(* IEC 61131-3 sources: Lasal-MCP/examples/SampleSource/LASALScreenAdvancedSolution/LASALScreenAdvancedSolution/LASALScreenAdvacnedSolution/Stations/Terminal/HMI/Class/MyFirstMyIO, 1 file *)

(* ---- MyFirstMyIO.st ---- *)
(*!
<Class
	Name               = "MyFirstMyIO"
	Revision           = "0.0"
	RealtimeTask       = "false"
	CyclicTask         = "false"
	BackgroundTask     = "false"
	Sigmatek           = "false"
	OSInterface        = "false"
	HighPriority       = "false"
	Automatic          = "false"
	UpdateMode         = "Prescan"
	SharedCommandTable = "true"
	Objectsize         = "(450,180)">
	<Channels>
		<Server Name="Number" Visualized="false" Initialize="false" WriteProtected="true" Retentive="false"/>
		<Client Name="_Grafix" Required="false" Internal="false"/>
	</Channels>
	<Network Name="MyFirstMyIO">
		<!-- List of Components in this network -->
		<Components>
			<Object
				Name       = "_base"
				Class      = "_MyIO"
				Position   = "(218,120)"
				Visualized = "true"
				Remotely   = "true">
				<Channels>
					<Server Name="Refresh"/>
					<Server Name="Server0"/>
					<Client Name="Graphic"/>
					<Client Name="Lse"/>
				</Channels>
			</Object>
		</Components>
		<Comments>
		</Comments>
		<!-- List of Connections in this network -->
		<Connections>
			<Connection Source="this.Server0" Destination="_base.Server0" Vertices="(706,210),(534,210),"/>
			<Connection Source="this.Refresh" Destination="_base.Refresh" Vertices="(706,270),(534,270),"/>
			<Connection Source="_base.Lse" Destination="this.Lse" Vertices="(218,210),(38,210),"/>
		</Connections>
		<!-- Headerfiles -->
		<Options>
		</Options>
	</Network>
</Class>
*)
#pragma using _MyIO

MyFirstMyIO : CLASS
: _MyIO
  //Servers:
	Number 	: SvrCh_DINT;
  //Clients:
	_Grafix 	: CltChCmd__Grafix;
  //Variables:
  //Functions:
				//! <Function Comment="this method is called everytime when system wants to redraw the io" Name="Draw"/>
	FUNCTION __CDECL VIRTUAL GLOBAL Draw
		VAR_INPUT
			pio 	: ^_IO;			//! <Variable Comment="pointer to _IO information" Name="Draw.pio"/>
			pr 	: ^_RESULT;			//! <Variable Comment="pointer to _RESULT information" Name="Draw.pr"/>
			pv 	: ^_VARIABLE;			//! <Variable Comment="pointer to io _VARIABLE information" Name="Draw.pv"/>
			input 	: BOOL;			//! <Variable Comment="TRUE it&apos;s an input&#13;&#10;FALSE it&apos;s an output" Name="Draw.input"/>
		END_VAR
		VAR_OUTPUT
			retcode (EAX) 	: _DOIT;			//! <Variable Comment="for the returnstatement there are 3 different possibilities&#13;&#10;  _IDLE ..... the system should goon like it is (system goes on)&#13;&#10;  _IDIDIT ... i did it (system is ready)&#13;&#10;  _IFAILED .. i tried to do my best, but i failed (system is re" Name="Draw.retcode"/>
		END_VAR;
				//! <Function Comment="method is called cyclic during object is on screen&#13;&#10;&#13;&#10;pio ....... &#13;&#10;input .... TRUE it&apos;s an input / FALSE it&apos;s an output&#13;&#10;" Name="IF_Run"/>
	FUNCTION __CDECL VIRTUAL GLOBAL IF_Run
		VAR_INPUT
			pio 	: ^_IO;			//! <Variable Comment="pointer to _IO information given by LSE" Name="IF_Run.pio"/>
			input 	: BOOL;			//! <Variable Comment="TRUE it&apos;s an input&#13;&#10;FALSE it&apos;s an output" Name="IF_Run.input"/>
		END_VAR;
				//! <Function Comment="this method is called right away before the object will be destroyed.&#13;&#10;for example close picture or window&#13;&#10;" Name="IF_End"/>
	FUNCTION __CDECL VIRTUAL GLOBAL IF_End;
  //Tables:
	FUNCTION @STD
		VAR_OUTPUT
			ret_code	: CONFSTATES;
		END_VAR;
	FUNCTION GLOBAL TAB @CT_;
END_CLASS;

#pragma usingLtd _Grafix

FUNCTION __CDECL VIRTUAL GLOBAL MyFirstMyIO::Draw
  #pragma warning(disable:73);
  VAR_INPUT
    pio 	: ^_IO;
    pr 	: ^_RESULT;
    pv 	: ^_VARIABLE;
    input 	: BOOL;
  END_VAR
  #pragma warning(default:73);
  VAR_OUTPUT
    retcode (EAX) 	: _DOIT;
  END_VAR
  VAR
    act : _NEWSCREEN;
    txt : array[0..10] of char;
  END_VAR

  // Switch active screen to Off-Screen
  push_screen(p0:= #act);

  // Copy content to Off-Screen
  _Grafix.PutImage(image:= #pio^.image, x0:= DEFKOORD, y0:= DEFKOORD);

  // Draw frame for _MyIo area with Lines
  _Grafix.Line(x0:= pio^.space.xy1.x,
               y0:= pio^.space.xy1.y,
               x1:= pio^.space.xy2.x,
               y1:= pio^.space.xy1.y,
               attrib:= pio^.attrib,
               color:= pio^.coltxt);

  _Grafix.Line(x0:= pio^.space.xy2.x,
               y0:= pio^.space.xy1.y,
               x1:= pio^.space.xy2.x,
               y1:= pio^.space.xy2.y,
               attrib:= pio^.attrib,
               color:= pio^.coltxt);

  _Grafix.Line(x0:= pio^.space.xy2.x,
               y0:= pio^.space.xy2.y,
               x1:= pio^.space.xy1.x,
               y1:= pio^.space.xy2.y,
               attrib:= pio^.attrib,
               color:= pio^.coltxt);

  _Grafix.Line(x0:= pio^.space.xy1.x,
               y0:= pio^.space.xy2.y,
               x1:= pio^.space.xy1.x,
               y1:= pio^.space.xy1.y,
               attrib:= pio^.attrib,
               color:= pio^.coltxt);

  // Set Text to defined coords
  _Grafix.OutTextXY(x0:= pio^.space.xy1.x + 100,
                    y0:= pio^.space.xy1.y + 50,
                    textptr:= "My Text!",
                    attrib:= pio^.attrib,
                    color:= _Grafix.MakeColor(backcolor:= INVISIBLE, frontcolor:= WHITE),
                    chr_size:= sizeof(_ASCII));

  // Convert Number to CHAR
  DToA(p0:= #txt[0],
       x1:= Number,
       x2:= 16#0800,
       x3:= sizeof(_ASCII));

  // Set Text to defined space
  OutTextAlign(p0:= #txt[0],         // Pointer to the text
               x1:= 0,               // No fill characters
               p1:= #pio^.space,     // Pointer to the coords
               x2:= pio^.font,       // The font to be used
               x3:= pio^.attrib,     // Attributes to display
               x9:= pio^.frametype,  // Frame type
               x4:= pio^.coltxt,     // Text color
               x5:= _Grafix.MakeColor(backcolor:= INVISIBLE, frontcolor:= INVISIBLE), // Background color
               x6:= _Grafix.MakeColor(backcolor:= INVISIBLE, frontcolor:= INVISIBLE), // Foreground color
               x7:= sizeof(_ASCII));  // ASCII or UNI

  // Switch active screen to output
  pop_screen(p0:= #act);

  // copy Off-Screen to output
  copy_screen(p0:= #act, p1:= #pio^.space);

  retcode := _IDIDIT;

END_FUNCTION

FUNCTION __CDECL VIRTUAL GLOBAL MyFirstMyIO::IF_Run
  #pragma warning(disable:73);
	VAR_INPUT
		pio 	: ^_IO;
		input 	: BOOL;
	END_VAR
  #pragma warning(default:73);

  Number += 1;
  Refresh := 1;

END_FUNCTION

FUNCTION __CDECL VIRTUAL GLOBAL MyFirstMyIO::IF_End

  Number := 0;

END_FUNCTION
